{attribute 'qualified_only'}
{attribute 'strict'}
{attribute 'to_string'}
TYPE E_Sint :
(
	eOptionA := 0,
	eOptionB,
	eOptionC
) SINT;
END_TYPE

(* stored: Version 1.1.0.1, ProductVersion 3.1.4026.19
   DUT E_Sint: Id {eca89de3-6da3-4462-870b-c7a5273878b0} *)
